(* IEC 61131-3 sources: codesys-framework/txt/application/WeVe Core (library)/30 Module/FB_Module/Commands, 4 files *)

(* ---- CommandResult.method.st ---- *)
// Resultaat van een commando opvragen zonder iets te starten (fire-and-forget opvolgen).
// Blijft staan tot er een nieuw commando start. Idle = dit commando is niet het laatste.
//   40 : Await(fbGripper.CommandResult(E_GripperCmd.Open), iNext := 50, iOnError := 900, iState := _iState);
METHOD CommandResult : E_CommandResult
VAR_INPUT
	iCmd 		: INT;
END_VAR

// --- BEGIN IMPLEMENTATION ---

CommandResult := _fbCmd.ResultOf(iCmd := iCmd);

(* ---- CommandTimeoutEvent.method.st ---- *)
// Overschrijven als de module een event wil bij een commando-timeout:
// geef de index van dat event in de enum van de module terug.
//   METHOD PROTECTED CommandTimeoutEvent : INT
//   CommandTimeoutEvent := E_GripperEvents.CommandTimeout;
// In ConfigureEvents van de groep:
//   Configure(iEvent := E_GripperEvents.CommandTimeout, udiEventId := cEv_ModuleCommandTimeout,
//             eEventLevel := E_EventLevels.EventIsAlarm_OperatorLevel, xResetable := TRUE, sMessage := 'Command %0 timed out.');
// -1 = geen event (standaard).
METHOD PROTECTED CommandTimeoutEvent : INT
VAR_INPUT
END_VAR

// --- BEGIN IMPLEMENTATION ---

CommandTimeoutEvent := -1;

(* ---- ExecuteCommand.method.st ---- *)
// Door de afgeleide module overschrijven: elke cyclus in Execute aangeroepen met het actieve commando.
//   CASE iCmd OF
//       E_GripperCmd.Open  : ... IF _fbHw.IsOpen THEN _fbCmd.Finish(); END_IF
//       E_GripperCmd.Close : ...
//   END_CASE
// Klaar: _fbCmd.Finish(). Gefaald: _fbCmd.Fail() en de oorzaak melden via een event.
METHOD PROTECTED ExecuteCommand
VAR_INPUT
	iCmd 		: INT;
END_VAR

// --- BEGIN IMPLEMENTATION ---

// Basis kent geen commando's
_fbCmd.Fail();

(* ---- InvokeCommand.method.st ---- *)
// Door de publieke commando-methodes van de afgeleide module.
// Start het commando als de module klaar is (Standby), of geeft de status terug als het al loopt.
// Bij de start gaat de module naar Execute; xStart is dan 1 cyclus TRUE: neem de parameters over.
METHOD PROTECTED InvokeCommand : E_CommandResult
VAR_INPUT
	iCmd 		: INT;				// commando-id uit de enum van de module, > 0
	tTimeout 	: TIME := T#0S;		// max duur van het commando, T#0S = geen timeout
END_VAR
VAR_OUTPUT
	xStart 		: BOOL;
END_VAR

// --- BEGIN IMPLEMENTATION ---

InvokeCommand := _fbCmd.Invoke(
	iCmd 		:= iCmd,
	xAllowed 	:= _eState = E_ModuleStates.Standby OR _eState = E_ModuleStates.Execute,
	tTimeout 	:= tTimeout,
	xStart 		=> xStart);

IF xStart THEN
	_eState := E_ModuleStates.Execute;
END_IF
